(* IEC 61131-3 sources: plc-st-coding-agent/progress/evidence/v13_rescore_20261108/candidates/custom_minimax-m27, 22 files *)

(* ---- public-easy-02.st ---- *)
FUNCTION_BLOCK FB
VAR_INPUT
    value   : DWORD;
END_VAR

VAR_OUTPUT
    hasChanged      : BOOL;
    hasRisingEdges  : BOOL;
    risingBits      : DWORD;
    noOfRisingBits  : USINT;
    hasFallingEdges : BOOL;
    fallingBits     : DWORD;
    noOfFallingBits : USINT;
END_VAR

VAR
    prevValue : DWORD;
    i         : USINT;
    bitMask   : DWORD;
END_VAR

(* Detect edges *)
risingBits  := value AND NOT prevValue;
fallingBits := prevValue AND NOT value;
hasChanged  := (value <> prevValue);
hasRisingEdges  := (risingBits <> 0);
hasFallingEdges := (fallingBits <> 0);

(* Count set bits *)
noOfRisingBits  := 0;
noOfFallingBits := 0;
FOR i := 0 TO 31 DO
    bitMask := SHL(DWORD#1, i);
    IF (risingBits AND bitMask) <> 0 THEN
        noOfRisingBits := noOfRisingBits + 1;
    END_IF
    IF (fallingBits AND bitMask) <> 0 THEN
        noOfFallingBits := noOfFallingBits + 1;
    END_IF
END_FOR

(* Update history *)
prevValue := value;

END_FUNCTION_BLOCK

(* ---- public-easy-03.st ---- *)
FUNCTION_BLOCK FB
VAR_INPUT
    Value       : REAL;
    hiLevel     : REAL;
    loLevel     : REAL;
    hystWindow  : REAL;
END_VAR
VAR_OUTPUT
    hiAlarm : BOOL := FALSE;
    loAlarm : BOOL := FALSE;
    error   : BOOL := FALSE;
    status  : WORD := 0;
END_VAR

error := FALSE;
status := 0;

IF loLevel >= hiLevel THEN
    error := TRUE;
    status := 16#8001;
    hiAlarm := FALSE;
    loAlarm := FALSE;
    RETURN;
END_IF

IF hystWindow >= (hiLevel - loLevel) THEN
    error := TRUE;
    status := 16#8002;
    hiAlarm := FALSE;
    loAlarm := FALSE;
    RETURN;
END_IF

IF Value > hiLevel THEN
    hiAlarm := TRUE;
ELSIF Value < (hiLevel - hystWindow) THEN
    hiAlarm := FALSE;
END_IF

IF Value < loLevel THEN
    loAlarm := TRUE;
ELSIF Value > (loLevel + hystWindow) THEN
    loAlarm := FALSE;
END_IF

END_FUNCTION_BLOCK

(* ---- public-easy-04.st ---- *)
FUNCTION_BLOCK FB
VAR_INPUT
    VISCOSITY_OK      : BOOL;
    PASTE_E_STOP_NC   : BOOL;
    DebounceTime      : TIME;
    CycleTime         : TIME;
END_VAR

VAR_OUTPUT
    VFD_RUN           : BOOL;
    PUMP_MAINT_DUE    : BOOL;
    PUMP_RUNTIME_ACC  : LINT;
END_VAR

VAR
    debounceTimer : TON;
    firstScan     : BOOL := TRUE;
END_VAR

// Power‑up initialisation
IF firstScan THEN
    VFD_RUN          := FALSE;
    PUMP_RUNTIME_ACC := 0;
    PUMP_MAINT_DUE   := FALSE;
    debounceTimer(IN := FALSE, PT := DebounceTime);
    firstScan := FALSE;
ELSE
    // Debounce the viscosity signal – timer resets when ESTOP opens
    debounceTimer(IN := VISCOSITY_OK AND PASTE_E_STOP_NC, PT := DebounceTime);

    // Run command requires ESTOP closed and viscosity condition validated
    VFD_RUN := PASTE_E_STOP_NC AND debounceTimer.Q;

    // Accumulate runtime while the pump is actually running
    IF VFD_RUN THEN
        PUMP_RUNTIME_ACC := PUMP_RUNTIME_ACC + CycleTime; // TIME converts to ms
    END_IF;

    // Maintenance due after 500 h (500 h = 500·3600·1000 ms)
    PUMP_MAINT_DUE := (PUMP_RUNTIME_ACC >= LINT#500 * 3600 * 1000);
END_IF

END_FUNCTION_BLOCK

(* ---- public-easy-06.st ---- *)
FUNCTION_BLOCK FB
VAR_INPUT
    DO_LOW            : BOOL;
    AERATION_E_STOP_NC: BOOL;
END_VAR
VAR_OUTPUT
    BLOWER_RUN                 : BOOL;
    AERATION_BLOWER_CYCLE_COUNT: UINT;
END_VAR
VAR
    StartDelayCounter : UINT;
    PrevBlowerRun     : BOOL;
END_VAR

IF NOT AERATION_E_STOP_NC OR NOT DO_LOW THEN
    BLOWER_RUN := FALSE;
    StartDelayCounter := 0;
ELSIF StartDelayCounter < 5 THEN
    StartDelayCounter := StartDelayCounter + 1;
    BLOWER_RUN := FALSE;
ELSE
    BLOWER_RUN := TRUE;
END_IF

IF BLOWER_RUN AND NOT PrevBlowerRun THEN
    AERATION_BLOWER_CYCLE_COUNT := AERATION_BLOWER_CYCLE_COUNT + 1;
END_IF

PrevBlowerRun := BLOWER_RUN;

END_FUNCTION_BLOCK

(* ---- public-hard-01.st ---- *)
FUNCTION_BLOCK FB
VAR_INPUT
    estop            : BOOL;
    opeMode          : BOOL;
    valveAStart      : BOOL;
    valveBStart      : BOOL;
    valveCStart      : BOOL;
    valveDStart      : BOOL;
    mixMotorStart    : BOOL;
    autoStart        : BOOL;
    processMode      : BOOL;
    levelSensor      : INT;
    mixMotorComplete : BOOL;
END_VAR
VAR_OUTPUT
    valveARun    : BOOL;
    valveBRun    : BOOL;
    valveCRun    : BOOL;
    valveDRun    : BOOL;
    mixMotorRun  : BOOL;
END_VAR
VAR
    autoState         : INT := 0;
    prevValveAStart   : BOOL := FALSE;
    prevValveBStart   : BOOL := FALSE;
    prevValveCStart   : BOOL := FALSE;
    prevValveDStart   : BOOL := FALSE;
    prevMixMotorStart : BOOL := FALSE;
    prevAutoStart     : BOOL := FALSE;
    prevMixMotorComplete : BOOL := FALSE;
END_VAR

    // Emergency stop: highest priority, stop all equipment immediately
    IF NOT estop THEN
        valveARun   := FALSE;
        valveBRun   := FALSE;
        valveCRun   := FALSE;
        valveDRun   := FALSE;
        mixMotorRun := FALSE;
        autoState   := 0;
        prevAutoStart            := autoStart;
        prevMixMotorComplete     := mixMotorComplete;
        prevValveAStart          := valveAStart;
        prevValveBStart          := valveBStart;
        prevValveCStart          := valveCStart;
        prevValveDStart          := valveDStart;
        prevMixMotorStart        := mixMotorStart;
    ELSE
        // Mode transition reset
        IF opeMode THEN
            IF prevValveAStart OR prevValveBStart OR prevValveCStart OR prevValveDStart OR prevMixMotorStart THEN
                autoState := 0;
            END_IF
            prevValveAStart   := FALSE;
            prevValveBStart   := FALSE;
            prevValveCStart   := FALSE;
            prevValveDStart   := FALSE;
            prevMixMotorStart := FALSE;
        ELSE
            // Manual mode: rising edge toggles
            IF valveAStart AND NOT prevValveAStart THEN
                valveARun := NOT valveARun;
            END_IF;
            IF valveBStart AND NOT prevValveBStart THEN
                valveBRun := NOT valveBRun;
            END_IF;
            IF valveCStart AND NOT prevValveCStart THEN
                valveCRun := NOT valveCRun;
            END_IF;
            IF valveDStart AND NOT prevValveDStart THEN
                valveDRun := NOT valveDRun;
            END_IF;
            IF mixMotorStart AND NOT prevMixMotorStart THEN
                mixMotorRun := NOT mixMotorRun;
            END_IF;
        END_IF

        // Automatic mode state machine
        IF opeMode THEN
            // State 0: Idle, wait for autoStart rising edge
            IF autoState = 0 THEN
                valveARun   := FALSE;
                valveBRun   := FALSE;
                valveCRun   := FALSE;
                valveDRun   := FALSE;
                mixMotorRun := FALSE;
                IF autoStart AND NOT prevAutoStart THEN
                    autoState := 1;
                END_IF;

            // State 1: Fill with valve A
            ELSIF autoState = 1 THEN
                valveBRun   := FALSE;
                valveCRun   := FALSE;
                valveDRun   := FALSE;
                mixMotorRun := FALSE;
                IF levelSensor >= 50 THEN
                    valveARun := FALSE;
                    autoState := 2;
                ELSE
                    valveARun := TRUE;
                END_IF;

            // State 2: Fill with valve B
            ELSIF autoState = 2 THEN
                valveARun   := FALSE;
                valveCRun   := FALSE;
                valveDRun   := FALSE;
                mixMotorRun := FALSE;
                IF levelSensor >= 80 THEN
                    valveBRun := FALSE;
                    IF processMode THEN
                        autoState := 3;
                    ELSE
                        autoState := 4;
                    END_IF;
                ELSE
                    valveBRun := TRUE;
                END_IF;

            // State 3: Fill with valve C (processMode = true)
            ELSIF autoState = 3 THEN
                valveARun   := FALSE;
                valveBRun   := FALSE;
                valveDRun   := FALSE;
                mixMotorRun := FALSE;
                IF levelSensor >= 100 THEN
                    valveCRun := FALSE;
                    autoState := 4;
                ELSE
                    valveCRun := TRUE;
                END_IF;

            // State 4: Mixing
            ELSIF autoState = 4 THEN
                valveARun   := FALSE;
                valveBRun   := FALSE;
                valveCRun   := FALSE;
                valveDRun   := FALSE;
                mixMotorRun := TRUE;
                IF mixMotorComplete AND NOT prevMixMotorComplete THEN
                    mixMotorRun := FALSE;
                    valveDRun   := TRUE;
                    autoState   := 5;
                END_IF;

            // State 5: Discharge complete, wait for next autoStart
            ELSIF autoState = 5 THEN
                valveARun   := FALSE;
                valveBRun   := FALSE;
                valveCRun   := FALSE;
                mixMotorRun := FALSE;
                valveDRun   := TRUE;
                IF autoStart AND NOT prevAutoStart THEN
                    valveDRun := FALSE;
                    autoState := 0;
                END_IF;
            END_IF;
        END_IF;
    END_IF;

    // Update edge detection history
    prevValveAStart   := valveAStart;
    prevValveBStart   := valveBStart;
    prevValveCStart   := valveCStart;
    prevValveDStart   := valveDStart;
    prevMixMotorStart := mixMotorStart;
    prevAutoStart     := autoStart;
    prevMixMotorComplete := mixMotorComplete;

END_FUNCTION_BLOCK

(* ---- public-hard-03.st ---- *)
TYPE ST_Recipe :
STRUCT
    recipeID : INT;
    ingredientType : INT;
    ingredientRatio : REAL;
    productionTemperature : REAL;
END_STRUCT
END_TYPE

FUNCTION_BLOCK FB
VAR_INPUT
    addRecipe : BOOL;
    deleteRecipe : BOOL;
    modifyRecipe : BOOL;
    queryRecipe : BOOL;
    recipeIn : ST_Recipe;
END_VAR

VAR_OUTPUT
    recipeAdded : BOOL;
    recipeDeleted : BOOL;
    recipeModified : BOOL;
    recipeQueryResult : ST_Recipe;
    error : BOOL;
    status : WORD;
END_VAR

VAR_IN_OUT
    recipe : ARRAY[1..10] OF ST_Recipe;
END_VAR

VAR
    addRecipe_prev : BOOL;
    deleteRecipe_prev : BOOL;
    modifyRecipe_prev : BOOL;
    queryRecipe_prev : BOOL;
END_VAR

VAR_TEMP
    idx : INT;
    foundIdx : INT;
    emptyIdx : INT;
    isFound : BOOL;
    hasEmpty : BOOL;
END_VAR

    recipeAdded := FALSE;
    recipeDeleted := FALSE;
    recipeModified := FALSE;
    error := FALSE;
    status := 16#0000;

    IF addRecipe AND NOT addRecipe_prev THEN
        isFound := FALSE;
        FOR idx := 1 TO 10 DO
            IF recipe[idx].recipeID = recipeIn.recipeID AND recipeIn.recipeID <> 0 THEN
                isFound := TRUE;
                EXIT;
            END_IF
        END_FOR

        IF isFound THEN
            error := TRUE;
            status := 16#8002;
        ELSE
            hasEmpty := FALSE;
            emptyIdx := 0;
            FOR idx := 1 TO 10 DO
                IF recipe[idx].recipeID = 0 THEN
                    hasEmpty := TRUE;
                    emptyIdx := idx;
                    EXIT;
                END_IF
            END_FOR

            IF hasEmpty THEN
                recipe[emptyIdx] := recipeIn;
                error := FALSE;
                status := 16#0000;
                recipeAdded := TRUE;
            ELSE
                error := TRUE;
                status := 16#8003;
            END_IF
        END_IF;

    ELSIF deleteRecipe AND NOT deleteRecipe_prev THEN
        isFound := FALSE;
        foundIdx := 0;
        FOR idx := 1 TO 10 DO
            IF recipe[idx].recipeID = recipeIn.recipeID AND recipeIn.recipeID <> 0 THEN
                isFound := TRUE;
                foundIdx := idx;
                EXIT;
            END_IF
        END_FOR

        IF isFound THEN
            recipe[foundIdx].recipeID := 0;
            recipe[foundIdx].ingredientType := 0;
            recipe[foundIdx].ingredientRatio := 0.0;
            recipe[foundIdx].productionTemperature := 0.0;
            error := FALSE;
            status := 16#0000;
            recipeDeleted := TRUE;
        ELSE
            error := TRUE;
            status := 16#8004;
        END_IF;

    ELSIF modifyRecipe AND NOT modifyRecipe_prev THEN
        isFound := FALSE;
        foundIdx := 0;
        FOR idx := 1 TO 10 DO
            IF recipe[idx].recipeID = recipeIn.recipeID AND recipeIn.recipeID <> 0 THEN
                isFound := TRUE;
                foundIdx := idx;
                EXIT;
            END_IF
        END_FOR

        IF isFound THEN
            recipe[foundIdx] := recipeIn;
            error := FALSE;
            status := 16#0000;
            recipeModified := TRUE;
        ELSE
            error := TRUE;
            status := 16#8005;
        END_IF;

    ELSIF queryRecipe AND NOT queryRecipe_prev THEN
        isFound := FALSE;
        foundIdx := 0;
        FOR idx := 1 TO 10 DO
            IF recipe[idx].recipeID = recipeIn.recipeID AND recipeIn.recipeID <> 0 THEN
                isFound := TRUE;
                foundIdx := idx;
                EXIT;
            END_IF
        END_FOR

        IF isFound THEN
            recipeQueryResult := recipe[foundIdx];
            error := FALSE;
            status := 16#0000;
        ELSE
            recipeQueryResult.recipeID := 0;
            recipeQueryResult.ingredientType := 0;
            recipeQueryResult.ingredientRatio := 0.0;
            recipeQueryResult.productionTemperature := 0.0;
            error := TRUE;
            status := 16#8001;
        END_IF;
    END_IF

    addRecipe_prev := addRecipe;
    deleteRecipe_prev := deleteRecipe;
    modifyRecipe_prev := modifyRecipe;
    queryRecipe_prev := queryRecipe;

END_FUNCTION_BLOCK

(* ---- public-medium-01.st ---- *)
TYPE ST_Pump :
STRUCT
    priority   : INT;
    selection  : BOOL;
    RunComd    : BOOL;
END_STRUCT
END_TYPE

FUNCTION_BLOCK FB
VAR_INPUT
    mode  : BOOL;
    start : BOOL;
    stop  : BOOL;
END_VAR
VAR_IN_OUT
    pumpGroup : ARRAY[1..5] OF ST_Pump;
END_VAR
VAR
    i         : INT;
    j         : INT;
    sortedIdx : ARRAY[1..5] OF INT;
    temp      : INT;
END_VAR

// sort pumps by priority (descending), stable on equal priority (lower index first)
sortedIdx[1] := 1;
sortedIdx[2] := 2;
sortedIdx[3] := 3;
sortedIdx[4] := 4;
sortedIdx[5] := 5;

FOR i := 1 TO 4 DO
    FOR j := i+1 TO 5 DO
        IF pumpGroup[sortedIdx[j]].priority > pumpGroup[sortedIdx[i]].priority THEN
            temp := sortedIdx[i];
            sortedIdx[i] := sortedIdx[j];
            sortedIdx[j] := temp;
        END_IF
    END_FOR
END_FOR

// stop has highest priority
IF stop THEN
    FOR i := 1 TO 5 DO
        pumpGroup[i].RunComd := FALSE;
    END_FOR
// start enables operation
ELSIF start THEN
    IF mode = FALSE THEN
        // Manual mode: selected pumps run
        FOR i := 1 TO 5 DO
            pumpGroup[i].RunComd := pumpGroup[i].selection;
        END_FOR
    ELSE
        // Automatic mode: top three priority pumps run
        FOR i := 1 TO 5 DO
            pumpGroup[i].RunComd := FALSE;
        END_FOR
        pumpGroup[sortedIdx[1]].RunComd := TRUE;
        pumpGroup[sortedIdx[2]].RunComd := TRUE;
        pumpGroup[sortedIdx[3]].RunComd := TRUE;
    END_IF
ELSE
    // start = FALSE -> no pump runs
    FOR i := 1 TO 5 DO
        pumpGroup[i].RunComd := FALSE;
    END_FOR
END_IF

END_FUNCTION_BLOCK

(* ---- public-medium-04.st ---- *)
FUNCTION_BLOCK FB
VAR_INPUT
    TemperatureSensorInput : REAL;
    SetTemperature : REAL;
END_VAR

VAR_OUTPUT
    CurrentTemperature : REAL;
    SetTempDisplay : REAL;
    HeaterStatus : BOOL;
    OverheatProtection : BOOL;
    HeaterOutput : BOOL;
END_VAR

VAR
    heating_time_count : INT := 0;
    overheat_wait_count : INT := 0;
    desired_heater : BOOL := FALSE;
    sensor_fault : BOOL := FALSE;
END_VAR

(* ---- Control logic ---- *)
sensor_fault := (TemperatureSensorInput < 0.0) OR (TemperatureSensorInput > 100.0);

desired_heater := FALSE;
IF NOT sensor_fault THEN
    IF TemperatureSensorInput < SetTemperature THEN
        desired_heater := TRUE;
    END_IF;
END_IF;

IF sensor_fault THEN
    HeaterOutput := FALSE;
    heating_time_count := 0;
    overheat_wait_count := 0;
    OverheatProtection := FALSE;
ELSE
    IF OverheatProtection THEN
        overheat_wait_count := overheat_wait_count + 1;
        HeaterOutput := FALSE;
        IF overheat_wait_count >= 3 THEN
            OverheatProtection := FALSE;
            overheat_wait_count := 0;
            heating_time_count := 0;
        END_IF;
    ELSE
        IF desired_heater THEN
            heating_time_count := heating_time_count + 1;
            IF heating_time_count > 5 THEN
                OverheatProtection := TRUE;
                HeaterOutput := FALSE;
                heating_time_count := 0;
                overheat_wait_count := 0;
            ELSE
                HeaterOutput := TRUE;
            END_IF;
        ELSE
            heating_time_count := 0;
            HeaterOutput := FALSE;
        END_IF;
    END_IF;
END_IF;

(* ---- Status outputs ---- *)
CurrentTemperature := TemperatureSensorInput;
SetTempDisplay := SetTemperature;
HeaterStatus := HeaterOutput;
END_FUNCTION_BLOCK

(* ---- public-medium-05.st ---- *)
TYPE StepEnum :
(
    Idle := 0,
    AtA,
    MovingAB,
    AtB,
    MovingBC,
    AtC
);
END_TYPE

FUNCTION_BLOCK FB
VAR_INPUT
    Mode            : BOOL;
    ForwardButton   : BOOL;
    ReverseButton   : BOOL;
    SensorA         : BOOL;
    SensorB         : BOOL;
    SensorC         : BOOL;
    ButtonA         : BOOL;
    ButtonB         : BOOL;
    ButtonC         : BOOL;
END_VAR
VAR_OUTPUT
    MotorForward    : BOOL;
    MotorReverse    : BOOL;
    CompletionLight : BOOL;
END_VAR
VAR
    prevMode            : BOOL := FALSE;
    prevForwardButton   : BOOL := FALSE;
    prevReverseButton   : BOOL := FALSE;
    prevButtonA         : BOOL := FALSE;
    prevButtonB         : BOOL := FALSE;
    prevButtonC         : BOOL := FALSE;
    prevSensorA         : BOOL := FALSE;
    prevSensorB         : BOOL := FALSE;
    prevSensorC         : BOOL := FALSE;
    currentStep         : StepEnum := Idle;
    buttonAPressed      : BOOL;
    buttonBPressed      : BOOL;
    buttonCPressed      : BOOL;
    sensorAArrived      : BOOL;
    sensorBArrived      : BOOL;
    sensorCArrived      : BOOL;
    sensorCRemoved      : BOOL;
END_VAR

// Detect mode change
IF Mode <> prevMode THEN
    IF NOT Mode THEN
        currentStep := Idle;
        CompletionLight := FALSE;
    END_IF;
END_IF;

// Compute edge detections
buttonAPressed   := ButtonA AND NOT prevButtonA;
buttonBPressed   := ButtonB AND NOT prevButtonB;
buttonCPressed   := ButtonC AND NOT prevButtonC;
sensorAArrived   := SensorA AND NOT prevSensorA;
sensorBArrived   := SensorB AND NOT prevSensorB;
sensorCArrived   := SensorC AND NOT prevSensorC;
sensorCRemoved   := prevSensorC AND NOT SensorC;

IF Mode = FALSE THEN
    // Manual mode
    MotorForward    := ForwardButton AND NOT ReverseButton;
    MotorReverse    := ReverseButton AND NOT ForwardButton;
    CompletionLight := FALSE;
ELSE
    // Automatic mode
    MotorReverse    := FALSE;
    MotorForward    := FALSE;

    CASE currentStep OF
        Idle:
            IF SensorA THEN
                currentStep := AtA;
            END_IF;

        AtA:
            IF buttonAPressed THEN
                currentStep := MovingAB;
                MotorForward := TRUE;
            END_IF;

        MovingAB:
            MotorForward := TRUE;
            IF sensorBArrived THEN
                MotorForward := FALSE;
                currentStep := AtB;
            END_IF;

        AtB:
            IF buttonBPressed THEN
                currentStep := MovingBC;
                MotorForward := TRUE;
            END_IF;

        MovingBC:
            MotorForward := TRUE;
            IF sensorCArrived THEN
                MotorForward := FALSE;
                currentStep := AtC;
            END_IF;

        AtC:
            IF buttonCPressed THEN
                CompletionLight := TRUE;
            END_IF;
            IF sensorCRemoved THEN
                CompletionLight := FALSE;
                currentStep := Idle;
            END_IF;
    END_CASE;
END_IF;

// Update previous inputs for next scan
prevMode            := Mode;
prevForwardButton   := ForwardButton;
prevReverseButton   := ReverseButton;
prevButtonA         := ButtonA;
prevButtonB         := ButtonB;
prevButtonC         := ButtonC;
prevSensorA         := SensorA;
prevSensorB         := SensorB;
prevSensorC         := SensorC;

END_FUNCTION_BLOCK

(* ---- public-medium-06.st ---- *)
FUNCTION_BLOCK FB
VAR_INPUT
    THICKNESS_FAULT        : BOOL;
    THICKNESS_SIGNAL_VALID : BOOL;
    CUTTING_RUN            : BOOL;
    FaultTimestamp         : DINT;
    CycleTime              : TIME;
END_VAR
VAR_OUTPUT
    THICKNESS_ALARM            : BOOL;
    Slab_Fault_Counter         : UINT;
    Slab_Runtime_Accumulator   : LINT;
    Slab_Fault_History         : ARRAY[0..4] OF DINT;
END_VAR
VAR
    FaultPrev       : BOOL := FALSE;
    AlarmHoldTimer  : TON;
END_VAR

(* Alarm control *)
IF NOT THICKNESS_SIGNAL_VALID THEN
    THICKNESS_ALARM      := FALSE;
    AlarmHoldTimer(IN := FALSE);
ELSE
    (* Rising edge of a valid fault *)
    IF THICKNESS_FAULT AND NOT FaultPrev THEN
        (* Increment fault counter *)
        Slab_Fault_Counter := Slab_Fault_Counter + 1;

        (* Shift history and store newest timestamp at index 0 *)
        Slab_Fault_History[4] := Slab_Fault_History[3];
        Slab_Fault_History[3] := Slab_Fault_History[2];
        Slab_Fault_History[2] := Slab_Fault_History[1];
        Slab_Fault_History[1] := Slab_Fault_History[0];
        Slab_Fault_History[0] := FaultTimestamp;

        (* Start 500 ms hold timer *)
        AlarmHoldTimer(IN := TRUE, PT := T#500ms);

        (* Activate alarm immediately *)
        THICKNESS_ALARM := TRUE;
    ELSE
        (* Normal alarm state handling *)
        IF THICKNESS_FAULT THEN
            (* Fault still present – keep alarm active *)
            THICKNESS_ALARM      := TRUE;
            AlarmHoldTimer(IN := TRUE, PT := T#500ms);
        ELSE
            (* Fault cleared – apply minimum hold period *)
            IF AlarmHoldTimer.Q THEN
                (* Hold time elapsed – deactivate alarm *)
                THICKNESS_ALARM      := FALSE;
                AlarmHoldTimer(IN := FALSE);
            ELSE
                (* Still within hold period *)
                THICKNESS_ALARM      := TRUE;
                AlarmHoldTimer(IN := TRUE, PT := T#500ms);
            END_IF
        END_IF
    END_IF
END_IF

(* Update edge detection variable *)
FaultPrev := THICKNESS_FAULT;

(* Runtime accumulation (only when signal valid, cutting running and no fault) *)
IF THICKNESS_SIGNAL_VALID AND CUTTING_RUN AND NOT THICKNESS_FAULT THEN
    Slab_Runtime_Accumulator := Slab_Runtime_Accumulator + (CycleTime / T#1ms);
END_IF

END_FUNCTION_BLOCK

(* ---- public-medium-07.st ---- *)
FUNCTION_BLOCK FB
VAR_INPUT
    OCCUPANCY_DETECTED : BOOL;
    ENERGY_SAVING_MODE : BOOL;
    HVAC_MODE_SELECTOR : INT;
END_VAR

VAR_OUTPUT
    SUPPLY_FAN_RUN : BOOL;
    TEMP_SETPOINT_ADJUST : INT;
END_VAR

VAR
    start_delay_timer : TON;
    delay_condition : BOOL;
    calculated_adjustment : INT;
END_VAR

SUPPLY_FAN_RUN := FALSE;
TEMP_SETPOINT_ADJUST := 0;

delay_condition := OCCUPANCY_DETECTED AND (HVAC_MODE_SELECTOR <> 3);

start_delay_timer(
    IN := delay_condition,
    PT := T#30s
);

IF delay_condition THEN
    SUPPLY_FAN_RUN := start_delay_timer.Q;
ELSE
    SUPPLY_FAN_RUN := FALSE;
END_IF;

CASE HVAC_MODE_SELECTOR OF
    0:
        IF OCCUPANCY_DETECTED THEN
            calculated_adjustment := 0;
        ELSE
            IF ENERGY_SAVING_MODE THEN
                calculated_adjustment := 3;
            ELSE
                calculated_adjustment := 2;
            END_IF;
        END_IF;

    1:
        IF OCCUPANCY_DETECTED THEN
            calculated_adjustment := 0;
        ELSE
            calculated_adjustment := 1;
        END_IF;

    2:
        IF OCCUPANCY_DETECTED THEN
            calculated_adjustment := 0;
        ELSE
            calculated_adjustment := 4;
        END_IF;

    3:
        calculated_adjustment := 4;

ELSE
    calculated_adjustment := 0;
END_CASE;

IF calculated_adjustment < -4 THEN
    TEMP_SETPOINT_ADJUST := -4;
ELSIF calculated_adjustment > 4 THEN
    TEMP_SETPOINT_ADJUST := 4;
ELSE
    TEMP_SETPOINT_ADJUST := calculated_adjustment;
END_IF;

END_FUNCTION_BLOCK

(* ---- public-medium-08.st ---- *)
FUNCTION_BLOCK FB
VAR_INPUT
    ipText: STRING(254);
END_VAR
VAR_OUTPUT
    ipValue: UDINT;
END_VAR
VAR
    len         : INT;
    pos         : INT;
    c           : CHAR;
    segCount    : INT;
    curVal      : UDINT;
    inSegment   : BOOL;
    segValues   : ARRAY[1..4] OF BYTE;
    ok          : BOOL;
END_VAR

// Reset outputs and internal state each cycle
ipValue   := 0;
ok        := TRUE;
segCount  := 0;
curVal    := 0;
inSegment := FALSE;

// Length of input string
len := LEN(ipText);
pos := 1;

// Parse characters
WHILE (pos <= len) AND ok DO
    c := ipText[pos];
    IF c = '.' THEN
        // End of current segment
        IF NOT inSegment THEN
            ok := FALSE;          // empty segment
            EXIT;
        END_IF
        // Store segment value
        segCount := segCount + 1;
        IF segCount > 4 THEN
            ok := FALSE;
            EXIT;
        END_IF
        segValues[segCount] := TO_BYTE(curVal);
        // Prepare for next segment
        curVal    := 0;
        inSegment := FALSE;
    ELSE
        // Expect decimal digit
        IF (c >= '0') AND (c <= '9') THEN
            curVal := curVal * 10 + UDINT(CHAR_TO_INT(c) - 48);
            IF curVal > 255 THEN
                ok := FALSE;
                EXIT;
            END_IF
            inSegment := TRUE;
        ELSE
            ok := FALSE;
            EXIT;
        END_IF
    END_IF
    pos := pos + 1;
END_WHILE

// Handle the last segment (if any)
IF ok THEN
    IF inSegment THEN
        segCount := segCount + 1;
        IF segCount > 4 THEN
            ok := FALSE;
        ELSE
            segValues[segCount] := TO_BYTE(curVal);
        END_IF
    ELSE
        // No digits after last dot or empty final segment
        ok := FALSE;
    END_IF
END_IF

// Assemble the 32‑bit address in network byte order
IF ok AND (segCount = 4) THEN
    ipValue := SHL(UDINT(segValues[1]), 24) OR
               SHL(UDINT(segValues[2]), 16) OR
               SHL(UDINT(segValues[3]), 8)  OR
               UDINT(segValues[4]);
ELSE
    ipValue := 0;
END_IF

END_FUNCTION_BLOCK

(* ---- self-easy-01.st ---- *)
FUNCTION_BLOCK FB
VAR_INPUT
    enable    : BOOL;
    values    : ARRAY[1..8] OF INT;
    count     : INT;
    avgEnable : BOOL;
END_VAR

VAR_OUTPUT
    avgOut : REAL;
END_VAR

VAR
    sumVal     : DINT;
    idx        : INT;
    validCnt   : INT;
END_VAR

// Default: keep previous output (no write occurs when conditions unmet)
// Guard: enable must be TRUE, avgEnable must be TRUE
IF enable AND avgEnable THEN
    // Guard: count must be positive (prevents div-by-zero per S1)
    IF count > 0 THEN
        // Clamp to array bound per requirement 3
        validCnt := count;
        IF validCnt > 8 THEN
            validCnt := 8;
        END_IF

        // Sum with DINT to avoid INT overflow
        sumVal := 0;
        FOR idx := 1 TO validCnt DO
            sumVal := sumVal + values[idx];
        END_FOR

        // Real division; validCnt > 0 guarantees no div-by-zero
        avgOut := DINT_TO_REAL(sumVal) / DINT_TO_REAL(validCnt);
    END_IF;
END_IF;

END_FUNCTION_BLOCK

(* ---- self-easy-02.st ---- *)
FUNCTION_BLOCK FB
VAR_INPUT
    tankLevel : REAL;
    outletFlow : REAL;
    inletPermit : BOOL;
    resetBtn : BOOL;
END_VAR
VAR_OUTPUT
    pumpRun : BOOL;
    alarmHigh : BOOL;
    alarmLow : BOOL;
    outletValveOpen : BOOL;
END_VAR
VAR
    lastResetBtn : BOOL := FALSE;
    internalAlarmHigh : BOOL := FALSE;
    internalAlarmLow : BOOL := FALSE;
    risingReset : BOOL;
END_VAR

risingReset := resetBtn AND NOT lastResetBtn;
lastResetBtn := resetBtn;

IF tankLevel >= 85.0 THEN
    internalAlarmHigh := TRUE;
ELSIF internalAlarmHigh AND risingReset AND (tankLevel < 85.0) THEN
    internalAlarmHigh := FALSE;
END_IF

IF tankLevel <= 15.0 THEN
    internalAlarmLow := TRUE;
ELSIF internalAlarmLow AND risingReset AND (tankLevel > 15.0) THEN
    internalAlarmLow := FALSE;
END_IF

IF internalAlarmHigh THEN
    pumpRun := FALSE;
ELSIF inletPermit AND (tankLevel < 85.0) AND (tankLevel >= 15.0) THEN
    pumpRun := TRUE;
ELSE
    pumpRun := FALSE;
END_IF

IF internalAlarmLow THEN
    outletValveOpen := FALSE;
ELSIF pumpRun THEN
    outletValveOpen := TRUE;
ELSE
    outletValveOpen := FALSE;
END_IF

alarmHigh := internalAlarmHigh;
alarmLow := internalAlarmLow;

END_FUNCTION_BLOCK

(* ---- self-hard-01.st ---- *)
FUNCTION_BLOCK FB
VAR_INPUT
    flowLow   : BOOL;
    ackBtn    : BOOL;
    sensorOK  : BOOL;
END_VAR
VAR_OUTPUT
    alarmActive : BOOL;
    alarmAcked  : BOOL;
    highHigh    : BOOL;
END_VAR
VAR
    prevAckBtn    : BOOL := FALSE;
    prevFlowLow   : BOOL := FALSE;
    xAlarmActive  : BOOL := FALSE;
    xAlarmAcked   : BOOL := FALSE;
END_VAR

(* New alarm on rising edge of flowLow *)
IF flowLow AND NOT prevFlowLow THEN
    xAlarmActive := TRUE;
    xAlarmAcked  := FALSE;
END_IF

(* Condition disappeared: set pending flag *)
IF NOT flowLow AND prevFlowLow THEN
    IF xAlarmActive AND NOT xAlarmAcked THEN
        xAlarmAcked := TRUE;
    END_IF;
END_IF

(* Acknowledge on rising edge of ack button *)
IF ackBtn AND NOT prevAckBtn THEN
    IF flowLow = FALSE AND xAlarmActive AND xAlarmAcked THEN
        xAlarmActive := FALSE;
        xAlarmAcked  := FALSE;
    ELSIF flowLow = TRUE AND xAlarmActive THEN
        xAlarmAcked := TRUE;
    END_IF;
END_IF

(* High‑priority alarm for sensor failure *)
highHigh := NOT sensorOK;

(* Drive outputs *)
alarmActive := xAlarmActive;
alarmAcked  := xAlarmAcked;

(* Update edge‑detection history *)
prevAckBtn  := ackBtn;
prevFlowLow := flowLow;

END_FUNCTION_BLOCK

(* ---- self-hard-02.st ---- *)
FUNCTION_BLOCK FB
VAR_INPUT
    startBtn    : BOOL;
    abortBtn    : BOOL;
    setpoint    : REAL;
    pv          : REAL;
    maxDuration : INT;
END_VAR
VAR_OUTPUT
    elapsed : INT;
    phase   : INT;
    timeout : BOOL;
END_VAR
VAR
    prevStartBtn : BOOL := FALSE;
    prevAbortBtn : BOOL := FALSE;
    risingStart  : BOOL;
END_VAR

(* Rising edge of start *)
risingStart := startBtn AND NOT prevStartBtn;

(* New start overrides abort to begin fresh batch *)
IF risingStart THEN
    elapsed := 0;
    timeout := FALSE;
    phase   := 1;
(* Abort has priority during normal operation (phases 1/2/3/0) *)
ELSIF abortBtn THEN
    phase := 9;
ELSE
    (* Normal operation *)
    IF phase = 1 THEN
        elapsed := elapsed + 1;
        IF pv >= setpoint THEN
            phase := 2;
        END_IF
    ELSIF phase = 2 THEN
        elapsed := elapsed + 1;
        IF elapsed >= maxDuration THEN
            timeout := TRUE;
            phase   := 3;
        END_IF
    END_IF
    (* Phases 0 and 3: wait for start *)
END_IF

(* Update edge‑detection history *)
prevStartBtn := startBtn;
prevAbortBtn := abortBtn;

END_FUNCTION_BLOCK

(* ---- self-hard-03.st ---- *)
FUNCTION_BLOCK FB
VAR_INPUT
    pushEn  : BOOL;
    pushItem: INT;
    popEn   : BOOL;
END_VAR

VAR_IN_OUT
    fifo : ARRAY[1..8] OF INT;
END_VAR

VAR_OUTPUT
    count : INT;
    full  : BOOL;
    empty : BOOL;
    head  : INT;
END_VAR

VAR
    prevPushEn : BOOL;
    prevPopEn  : BOOL;
    risingPush : BOOL;
    risingPop  : BOOL;
    i          : INT;
END_VAR

// Step 1: Rising edge detection
risingPush := pushEn AND NOT prevPushEn;
risingPop  := popEn  AND NOT prevPopEn;

// Step 2: Pop first when both edges occur in same cycle
IF risingPop THEN
    IF count > 0 THEN
        FOR i := 1 TO count - 1 DO
            fifo[i] := fifo[i + 1];
        END_FOR
        fifo[count] := 0;
        count := count - 1;
    END_IF
END_IF

// Step 3: Push after pop
IF risingPush THEN
    IF count < 8 THEN
        count := count + 1;
        fifo[count] := pushItem;
    END_IF
END_IF

// Step 4: Update outputs
empty := (count = 0);
full  := (count = 8);

IF count > 0 THEN
    head := fifo[1];
ELSE
    head := 0;
END_IF

// Step 5: Update edge history for next scan
prevPushEn := pushEn;
prevPopEn  := popEn;

END_FUNCTION_BLOCK

(* ---- self-hard-05.st ---- *)
FUNCTION_BLOCK FB
VAR_INPUT
    runRequest  : BOOL;
    flameOK     : BOOL;
    o2Valid     : BOOL;
    o2PV        : REAL;
    baseAir     : REAL;
    resetBtn    : BOOL;
END_VAR
VAR_OUTPUT
    fuelPermit  : BOOL;
    trimEnable  : BOOL;
    airTrim     : REAL;
    airCommand  : REAL;
    tripLatched : BOOL;
    o2Fault     : BOOL;
END_VAR
VAR
    prevResetBtn : BOOL := FALSE;
END_VAR

// S2: 跳闸置位与清除（清除需复位上升沿且 flameOK=FALSE 且 runRequest=FALSE）
IF prevResetBtn AND NOT resetBtn AND NOT runRequest AND NOT flameOK THEN
    tripLatched := FALSE;
ELSIF runRequest AND NOT flameOK THEN
    tripLatched := TRUE;
END_IF;

// 记录复位按钮上一状态（边沿检测）
prevResetBtn := resetBtn;

// o2Fault：独立于 tripLatched，只切除修正不切除燃料
o2Fault := NOT o2Valid OR o2PV < 0.0 OR o2PV > 21.0;

// fuelPermit：runRequest AND flameOK AND NOT tripLatched
fuelPermit := runRequest AND flameOK AND NOT tripLatched;

// trimEnable：fuelPermit AND NOT o2Fault
trimEnable := fuelPermit AND NOT o2Fault;

// airTrim 钳位 ±10；trimEnable=FALSE 时强制为 0.0
IF trimEnable THEN
    airTrim := 2.0 * (2.0 - o2PV);
    IF airTrim > 10.0 THEN
        airTrim := 10.0;
    ELSIF airTrim < -10.0 THEN
        airTrim := -10.0;
    END_IF;
ELSE
    airTrim := 0.0;
END_IF;

// airCommand：fuelPermit=FALSE 时强制为 0.0；否则钳位 0..100
IF NOT fuelPermit THEN
    airCommand := 0.0;
ELSE
    airCommand := baseAir + airTrim;
    IF airCommand > 100.0 THEN
        airCommand := 100.0;
    ELSIF airCommand < 0.0 THEN
        airCommand := 0.0;
    END_IF;
END_IF;
END_FUNCTION_BLOCK

(* ---- self-hard-06.st ---- *)
FUNCTION_BLOCK FB
VAR_INPUT
    runRequest : BOOL;
    pressure : REAL;
    pressureValid : BOOL;
    fuelFlow : REAL;
    steamFlow : REAL;
    outletCmd : INT;
    outletFeedback : INT;
    resetBtn : BOOL;
END_VAR
VAR_OUTPUT
    tripLatched : BOOL;
    fuelPermit : BOOL;
    currentCauseMask : WORD;
    latchedCauseMask : WORD;
    diagnosticActive : BOOL;
END_VAR
VAR
    tripLatchedState : BOOL := FALSE;
    resetBtnPrev : BOOL := FALSE;
    valveStuckCounter : INT := 0;
    latchedCauseMaskInternal : WORD := 0;
    tripCondition : BOOL;
    resetBtnRising : BOOL;
    tempMask : WORD;
END_VAR

// 检测复位按钮上升沿
resetBtnRising := resetBtn AND NOT resetBtnPrev;

// 判断跳闸条件
tripCondition := (runRequest AND pressureValid AND (pressure >= 4500.0)) OR (runRequest AND NOT pressureValid);

// 跳闸条件成立则置位自保持
IF tripCondition THEN
    tripLatchedState := TRUE;
END_IF

// 复位上升沿且满足清除条件时解除跳闸
IF resetBtnRising AND NOT runRequest AND pressureValid AND (pressure <= 4200.0) THEN
    tripLatchedState := FALSE;
    latchedCauseMaskInternal := 0; // 复位时清零故障记录
END_IF

// 更新阀门卡滞计数器（跨周期记忆）
IF runRequest THEN
    IF pressureValid AND (pressure >= 4500.0) AND (outletCmd >= 50) AND (outletFeedback <= 10) THEN
        valveStuckCounter := valveStuckCounter + 1;
    ELSE
        valveStuckCounter := 0;
    END_IF
ELSE
    valveStuckCounter := 0;
END_IF

// 计算本周期线索掩码
tempMask := 0;
IF NOT runRequest THEN
    tempMask := 0;
ELSE
    IF pressureValid AND (pressure < 4500.0) THEN
        tempMask := 0;
    ELSE
        // bit0: 变送器失效
        IF NOT pressureValid THEN
            tempMask := tempMask OR 1;
        END_IF
        // bit1: 减温减压阀卡滞（连续3拍及以上）
        IF valveStuckCounter >= 3 THEN
            tempMask := tempMask OR 2;
        END_IF
        // bit2: 燃烧过剩
        IF (fuelFlow >= 4.0) AND (steamFlow <= 10.0) THEN
            tempMask := tempMask OR 4;
        END_IF
        // bit3: 未定位
        IF (tempMask = 0) AND pressureValid AND (pressure >= 4500.0) THEN
            tempMask := tempMask OR 8;
        END_IF
    END_IF
END_IF

// 跳闸时按位或累积线索
IF tripLatchedState THEN
    latchedCauseMaskInternal := latchedCauseMaskInternal OR tempMask;
END_IF

// 更新历史变量
resetBtnPrev := resetBtn;

// 输出赋值
tripLatched := tripLatchedState;
fuelPermit := runRequest AND NOT tripLatchedState;
currentCauseMask := tempMask;
latchedCauseMask := latchedCauseMaskInternal;
diagnosticActive := (tempMask <> 0);

END_FUNCTION_BLOCK

(* ---- self-medium-02.st ---- *)
FUNCTION_BLOCK FB
VAR_INPUT
    enable      : BOOL;
    rawValue    : REAL;
END_VAR

VAR_OUTPUT
    filteredValue : REAL;
    windowFull    : BOOL;
    sampleCount   : INT;
END_VAR

VAR
    buffer       : ARRAY[0..7] OF REAL;
    writeIndex   : INT;
    sumValue     : REAL;
    index        : INT;
END_VAR

IF NOT enable THEN
    sampleCount := 0;
    windowFull := FALSE;
    writeIndex := 0;
    sumValue := 0.0;

    FOR index := 0 TO 7 DO
        buffer[index] := 0.0;
    END_FOR;
ELSE
    sumValue := 0.0;

    IF sampleCount < 8 THEN
        FOR index := 0 TO sampleCount - 1 DO
            sumValue := sumValue + buffer[index];
        END_FOR;

        sumValue := sumValue + rawValue;
        filteredValue := sumValue / INT_TO_REAL(sampleCount + 1);
    ELSE
        FOR index := 0 TO 7 DO
            sumValue := sumValue + buffer[index];
        END_FOR;

        sumValue := sumValue + rawValue - buffer[writeIndex];
        filteredValue := sumValue / 8.0;
    END_IF;

    buffer[writeIndex] := rawValue;

    IF writeIndex = 7 THEN
        writeIndex := 0;
    ELSE
        writeIndex := writeIndex + 1;
    END_IF;

    IF sampleCount < 8 THEN
        sampleCount := sampleCount + 1;
    END_IF;

    IF sampleCount >= 8 THEN
        windowFull := TRUE;
    END_IF;
END_IF

END_FUNCTION_BLOCK

(* ---- self-medium-03.st ---- *)
FUNCTION_BLOCK FB
VAR_INPUT
    openBtn    : BOOL;
    closeBtn   : BOOL;
    openLimit  : BOOL;
    closeLimit : BOOL;
    obstacle   : BOOL;
END_VAR

VAR_OUTPUT
    motorUp   : BOOL;
    motorDown : BOOL;
    errorFlag : BOOL;
END_VAR

VAR
    state        : INT := 0;   // 0=IDLE, 1=OPENING, 2=CLOSING, 3=FAULT
    prevOpenBtn  : BOOL := FALSE;
    prevCloseBtn : BOOL := FALSE;
END_VAR

VAR
    openRising  : BOOL;
    closeRising : BOOL;
END_VAR

// Detect rising edges of the push‑button inputs
openRising  := openBtn AND NOT prevOpenBtn;
closeRising := closeBtn AND NOT prevCloseBtn;

// Update button history for next scan
prevOpenBtn  := openBtn;
prevCloseBtn := closeBtn;

// ------------------------------------------------------------
// Finite State Machine
// ------------------------------------------------------------
CASE state OF
    // --------------------------------------------------------
    // IDLE – waiting for a command
    // --------------------------------------------------------
    0:
        motorUp   := FALSE;
        motorDown := FALSE;
        errorFlag := FALSE;

        IF openRising AND NOT openLimit THEN
            state := 1;               // start opening
        ELSIF closeRising AND NOT closeLimit THEN
            state := 2;               // start closing
        END_IF

    // --------------------------------------------------------
    // OPENING – motor raises the gate
    // --------------------------------------------------------
    1:
        motorUp   := TRUE;
        motorDown := FALSE;
        errorFlag := FALSE;

        IF openLimit THEN
            state := 0;               // reached open limit
        ELSIF obstacle THEN
            motorUp   := FALSE;       // stop motor immediately
            errorFlag := TRUE;
            state := 3;               // enter fault state
        END_IF

    // --------------------------------------------------------
    // CLOSING – motor lowers the gate
    // --------------------------------------------------------
    2:
        motorUp   := FALSE;
        motorDown := TRUE;
        errorFlag := FALSE;

        IF closeLimit THEN
            state := 0;               // reached close limit
        ELSIF obstacle THEN
            motorDown := FALSE;       // stop downward motion
            IF openLimit THEN
                // Already at open limit → just stop
                state := 0;
            ELSE
                motorUp := TRUE;      // reverse to opening
                state := 1;
            END_IF
        END_IF

    // --------------------------------------------------------
    // FAULT – motor stopped, error latched
    // --------------------------------------------------------
    3:
        motorUp   := FALSE;
        motorDown := FALSE;
        errorFlag := TRUE;

        // Reset allowed only when obstacle cleared and both buttons pressed (rising edges)
        IF (NOT obstacle) AND openRising AND closeRising THEN
            errorFlag := FALSE;
            state := 0;
        END_IF

END_CASE
END_FUNCTION_BLOCK

(* ---- self-medium-04.st ---- *)
FUNCTION_BLOCK FB
VAR_INPUT
    startBtn   : BOOL;
    resetBtn   : BOOL;
    doneSensor : BOOL;
    targetVol  : REAL;
    flowVol    : REAL;
END_VAR
VAR_OUTPUT
    valveOpen  : BOOL;
    fillsToday : INT;
END_VAR
VAR
    eState       : INT;     // 0=IDLE, 1=FILLING, 2=WAITING_CONFIRM
    accumulator  : REAL;
    lastStartBtn : BOOL;
    lastResetBtn : BOOL;
    risingStart  : BOOL;
    risingReset  : BOOL;
END_VAR

    // ---- Edge detection -------------------------------------------------
    risingStart := startBtn AND NOT lastStartBtn;
    risingReset := resetBtn AND NOT lastResetBtn;

    // ---- Reset handling (highest priority) -------------------------------
    IF risingReset THEN
        valveOpen   := FALSE;
        accumulator := 0.0;
        fillsToday  := 0;
        eState      := 0;    // IDLE
    ELSE
        // ---- State machine -----------------------------------------------
        CASE eState OF
            0:  // IDLE
                IF risingStart THEN
                    valveOpen   := TRUE;
                    accumulator := 0.0;
                    eState      := 1;  // FILLING
                ELSE
                    valveOpen := FALSE;
                END_IF

            1:  // FILLING
                accumulator := accumulator + flowVol;
                IF accumulator >= targetVol THEN
                    valveOpen := FALSE;
                    eState    := 2;    // WAITING_CONFIRM
                END_IF

            2:  // WAITING_CONFIRM
                valveOpen := FALSE;
                IF doneSensor THEN
                    fillsToday := fillsToday + 1;
                    eState     := 0;    // IDLE
                END_IF
        END_CASE
    END_IF

    // ---- Update edge histories --------------------------------------------
    lastStartBtn := startBtn;
    lastResetBtn := resetBtn;

END_FUNCTION_BLOCK
